// TIA Portal V20 export
FUNCTION_BLOCK "Melden_VisuAllgemein"   // FB127, LAD
{ S7_Optimized_Access := 'TRUE' }
// stored: MemoryReserve 100, SetENOAutomatically false
   VAR
      Register_leer : "Teile Status";
      auf_Seite_Richten { S7_SetPoint := 'True'} : Bool;
      Flanke_Bildwechsel { S7_SetPoint := 'True'} : R_TRIG;
      Bild_tmp { S7_SetPoint := 'True'} : DInt;
      WartezeitSicherung_Reset { S7_SetPoint := 'True'} : TON_TIME;
      Flanke_Türe8_schließen { S7_SetPoint := 'True'} : R_TRIG;
      Flanke_Türe8_öffnen { S7_SetPoint := 'True'} : R_TRIG;
   END_VAR
   VAR RETAIN
      Artikelnummer_tmp { ExternalAccessible := 'False'; ExternalVisible := 'False'; ExternalWritable := 'False'} : String;
   END_VAR
   VAR
      VZ_Leerfahren { S7_SetPoint := 'True'} : TON_TIME;
   END_VAR
   VAR_TEMP
      test : Bool;
   END_VAR
BEGIN

REGION Network 1 (SCL): Richten oder Einzelschrittseite aufgerufen
   CASE "HMI_SYS"."Aktueller Bildschirm" OF
       75:
           #auf_Seite_Richten := true;
       ELSE
           #auf_Seite_Richten := false;
   END_CASE;
END_REGION

REGION Network 2 (SCL): Artikel wurde gewechselt


   IF #Artikelnummer_tmp <> "HMI_COM".Artikelnummer_String THEN
       "HMI_COM".Artikel_gewechselt := true;
       #Artikelnummer_tmp := "HMI_COM".Artikelnummer_String;
   ELSIF "HMI_COM".Grundstellung_Gesamt AND  "HMI_COM".Artikel_gewechselt THEN

       "HMI_COM".Artikel_gewechselt := false;

   END_IF;
END_REGION

NETWORK
TITLE = Übergabe Anwahl Richten
      A     #auf_Seite_Richten;
      JC    m003;

      JU    m001;
m003: NOP   0;

      A     "03_Betriebsart_DB"."NOT-HALT OK";
      A     "03_Betriebsart_DB"."Schutztüren OK";
      JCN   m001;


      A     "HMI_COM".Richten_Gesamtanlage;
      JCN   m002;

      SET;
      S     "HMI_BETR_ART_POS".POS3_0.Taster_Anwahl_GS;


m002: NOP   0;

      A     "HMI_BETR_ART_POS".POS3_0.Taster_Anwahl_GS;
      S     "POS3_0_Signal".Station.SK_Freigabe_Richten;
      =     "POS3_0_Signal".Schrittkette.INIT_SQ;
      R     "HMI_BETR_ART_POS".POS3_0.Taster_Anwahl_GS;


      A     "HMI_COM".Richten_Gesamtanlage;
      R     "HMI_COM".Richten_Gesamtanlage;

m001: NOP   0;


NETWORK
TITLE = Tippbetrieb Aktiv
      A     "POS3_0_Signal".Schrittkette.AUTO_ON;


      =     "HMI_COM".Einzelschritt.Status_Anw;


NETWORK
TITLE = Antriebe sind Ein
      SET;

      =     "HMI_COM".Antriebe_sind_EIN;

REGION Network 6 (SCL): Übergabe Türen Not Halt
   // Allgemeine HMI Übergabe 

   "HMI_COM"."NOT-HALT_OK" := "03_Betriebsart_DB"."NOT-HALT OK";
   "HMI_COM".TUERE_OK := "03_Betriebsart_DB"."Schutztüren OK";




   // Übergabe welche Tür ist nicht verriegelt
   REGION Türen


       "HMI_COM".Tür_offen[1] := "DE_Rueckfuehrung_Tuer_1" AND ("03_Betriebsart_DB".BA_Automatik OR "03_Betriebsart_DB".BA_Manuell OR "03_Betriebsart_DB".BA_Richten);
       "HMI_COM".Tür_offen[2] := "DE_Rueckfuehrung_Tuer_2" AND ("03_Betriebsart_DB".BA_Automatik OR "03_Betriebsart_DB".BA_Manuell OR "03_Betriebsart_DB".BA_Richten);
    //   "HMI_COM".Tür_offen[3] := "DE_Rueckfuehrung_Tuer_3" AND ("03_Betriebsart_DB".BA_Automatik OR "03_Betriebsart_DB".BA_Manuell OR "03_Betriebsart_DB".BA_Richten);
    //   "HMI_COM".Tür_offen[4] := "DE_Rueckfuehrung_Tuer_4" AND ("03_Betriebsart_DB".BA_Automatik OR "03_Betriebsart_DB".BA_Manuell OR "03_Betriebsart_DB".BA_Richten);
    //   "HMI_COM".Tür_offen[5] := "DE_Rueckfuehrung_Tuer_5" AND ("03_Betriebsart_DB".BA_Automatik OR "03_Betriebsart_DB".BA_Manuell OR "03_Betriebsart_DB".BA_Richten);
    //   "HMI_COM".Tür_offen[6] := "DE_Rueckfuehrung_Tuer_6" AND ("03_Betriebsart_DB".BA_Automatik OR "03_Betriebsart_DB".BA_Manuell OR "03_Betriebsart_DB".BA_Richten);
    //   "HMI_COM".Tür_offen[7] := "DE2_0_Rückführung Tür 7" AND ("03_Betriebsart_DB".BA_Automatik OR "03_Betriebsart_DB".BA_Manuell OR "03_Betriebsart_DB".BA_Richten);
    //   "HMI_COM".Tür_offen[8] := "DE2_1_Rückführung Tür 8" AND ("03_Betriebsart_DB".BA_Automatik OR "03_Betriebsart_DB".BA_Manuell OR "03_Betriebsart_DB".BA_Richten);
    (*   "HMI_COM".Tür_offen[9] := "DE2_1_Rückführung Tür 8" AND ("03_Betriebsart_DB".BA_Automatik OR "03_Betriebsart_DB".BA_Manuell OR "03_Betriebsart_DB".BA_Richten);
       "HMI_COM".Tür_offen[10] := "DE2_1_Rückführung Tür 8" AND ("03_Betriebsart_DB".BA_Automatik OR "03_Betriebsart_DB".BA_Manuell OR "03_Betriebsart_DB".BA_Richten);
       "HMI_COM".Tür_offen[11] := "DE2_1_Rückführung Tür 8" AND ("03_Betriebsart_DB".BA_Automatik OR "03_Betriebsart_DB".BA_Manuell OR "03_Betriebsart_DB".BA_Richten);
       "HMI_COM".Tür_offen[12] := "DE2_1_Rückführung Tür 8" AND ("03_Betriebsart_DB".BA_Automatik OR "03_Betriebsart_DB".BA_Manuell OR "03_Betriebsart_DB".BA_Richten);
       "HMI_COM".Tür_offen[13] := "DE2_1_Rückführung Tür 8" AND ("03_Betriebsart_DB".BA_Automatik OR "03_Betriebsart_DB".BA_Manuell OR "03_Betriebsart_DB".BA_Richten);
       "HMI_COM".Tür_offen[14] := "DE2_1_Rückführung Tür 8" AND ("03_Betriebsart_DB".BA_Automatik OR "03_Betriebsart_DB".BA_Manuell OR "03_Betriebsart_DB".BA_Richten);
       "HMI_COM".Tür_offen[15] := "DE2_1_Rückführung Tür 8" AND ("03_Betriebsart_DB".BA_Automatik OR "03_Betriebsart_DB".BA_Manuell OR "03_Betriebsart_DB".BA_Richten); *)
    //   "HMI_COM".Tür_offen[16] := "DE2_1_Rückführung Tür 8" AND ("03_Betriebsart_DB".BA_Automatik OR "03_Betriebsart_DB".BA_Manuell OR "03_Betriebsart_DB".BA_Richten);

   END_REGION
END_REGION

REGION Network 7 (SCL): Rücksetzen der Stationen bei Grundbild



   #Flanke_Bildwechsel(CLK:="03_Betriebsart_DB".BA_Manuell AND #Bild_tmp <> "HMI_SYS"."Aktueller Bildschirm" );



   IF #Flanke_Bildwechsel.Q THEN

       #Bild_tmp := "HMI_SYS"."Aktueller Bildschirm";

    //IF ("HMI_SYS"."Aktueller Bildschirm" = 10125) OR ("03_Betriebsart_DB"."NOT-HALT OK" = false) THEN

       "HMI_COM".Manuell_Zylinder1.Status := 0;
       "HMI_COM".Manuell_Zylinder2.Status := 0;
       "HMI_COM".Manuell_Zylinder3.Status := 0;
       "HMI_COM".Manuell_Zylinder4.Status := 0;

       "HMI_COM".Manuell_Zylinder1.GS := FALSE;
       "HMI_COM".Manuell_Zylinder1.AS1 := FALSE;
       "HMI_COM".Manuell_Zylinder2.GS := FALSE;
       "HMI_COM".Manuell_Zylinder2.AS1 := FALSE;
       "HMI_COM".Manuell_Zylinder3.GS := FALSE;
       "HMI_COM".Manuell_Zylinder3.AS1 := FALSE;
       "HMI_COM".Manuell_Zylinder4.GS := FALSE;
       "HMI_COM".Manuell_Zylinder4.AS1 := FALSE;

      "HMI_COM".Manuell_Zylinder1.DA_GS := FALSE;
       "HMI_COM".Manuell_Zylinder1.DA_AS1 := FALSE;
       "HMI_COM".Manuell_Zylinder2.DA_GS := FALSE;
       "HMI_COM".Manuell_Zylinder2.DA_AS1 := FALSE;
       "HMI_COM".Manuell_Zylinder3.DA_GS := FALSE;
       "HMI_COM".Manuell_Zylinder3.DA_AS1 := FALSE;
       "HMI_COM".Manuell_Zylinder4.DA_GS := FALSE;
       "HMI_COM".Manuell_Zylinder4.DA_AS1 := FALSE;
     END_IF;
END_REGION

REGION Network 8 (SCL): Übertragung und Verwaltung Register



   "HMI_COM".Speichern_Register := false;
END_REGION

REGION Network 9 (SCL): Rucksetzen wenn Register nicht gelöscht
   IF (("HMI_SYS"."Aktueller Bildschirm" = 10001) OR ("HMI_SYS"."Aktueller Bildschirm" = 10010) OR ("HMI_SYS"."Aktueller Bildschirm" = 10020)
       OR ("HMI_SYS"."Aktueller Bildschirm" = 10030)) THEN

       "HMI_BETR_ART_POS".POS3_0.Taster_Reset_Teilestatus := FALSE;
       "HMI_BETR_ART_POS".POS3_1.Taster_Reset_Teilestatus := FALSE;
       "HMI_BETR_ART_POS".POS3_2.Taster_Reset_Teilestatus := FALSE;
       "HMI_BETR_ART_POS".POS3_3.Taster_Reset_Teilestatus := FALSE;
       "HMI_BETR_ART_POS".POS3_4.Taster_Reset_Teilestatus := FALSE;
       "HMI_BETR_ART_POS".POS4_0_Zuführung.Taster_Reset_Teilestatus := FALSE;
       "HMI_BETR_ART_POS".POS5_0_Zuführung.Taster_Reset_Teilestatus := FALSE;
       "HMI_BETR_ART_POS".POS5_0.Taster_Reset_Teilestatus := FALSE;
       "HMI_BETR_ART_POS".POS6_0.Taster_Reset_Teilestatus := FALSE;
       "HMI_BETR_ART_POS".POS7_0.Taster_Reset_Teilestatus := FALSE;
       "HMI_BETR_ART_POS".POS7_1.Taster_Reset_Teilestatus := FALSE;
       "HMI_BETR_ART_POS".POS7_2.Taster_Reset_Teilestatus := FALSE;
       "HMI_BETR_ART_POS".POS7_3.Taster_Reset_Teilestatus := FALSE;
       "HMI_BETR_ART_POS".POS7_4.Taster_Reset_Teilestatus := FALSE;
       "HMI_BETR_ART_POS".POS8_0.Taster_Reset_Teilestatus := FALSE;
       "HMI_BETR_ART_POS".POS9_0.Taster_Reset_Teilestatus := FALSE;
       "HMI_BETR_ART_POS".POS9_1.Taster_Reset_Teilestatus := FALSE;
       "HMI_BETR_ART_POS".POS9_2.Taster_Reset_Teilestatus := FALSE;
       "HMI_BETR_ART_POS".POS9_3.Taster_Reset_Teilestatus := FALSE;
       "HMI_BETR_ART_POS".POS9_4.Taster_Reset_Teilestatus := FALSE;
       "HMI_BETR_ART_POS".POS9_5.Taster_Reset_Teilestatus := FALSE;
       "HMI_BETR_ART_POS".POS9_6.Taster_Reset_Teilestatus := FALSE;
       "HMI_BETR_ART_POS".POS10_0.Taster_Reset_Teilestatus := FALSE;
       "HMI_BETR_ART_POS".POS11.Taster_Reset_Teilestatus := FALSE;
       "HMI_BETR_ART_POS".POS12.Taster_Reset_Teilestatus := FALSE;

   END_IF;
END_REGION

REGION Network 10 (SCL): Leerfahren
   "HMI_Signale".Leerfahren_angewaehlt := "HMI_COM".Leerfahren_angewaehlt;

   #VZ_Leerfahren(IN := "HMI_COM".Leerfahren_ende,
                  PT := t#3s);

   IF #VZ_Leerfahren.Q OR "HMI_COM".Leerfahren_angewaehlt = false THEN

       "HMI_COM".Leerfahren_ende := FALSE;
       "HMI_Signale".Leerfahren_ende := false;
       "HMI_COM".Leerfahren_angewaehlt := false;

       "HMI_COM".Leerfahren_laeuft := false; 
       "POS3_0_Signal".Station.SK_Freigabe_Auto := false;




   END_IF;
END_REGION

REGION Network 11 (SCL): Bildaufrufe


       // Bei Not-Aus Aufruf Grundbild
       IF "03_Betriebsart_DB".BA_0_FP = TRUE OR
           "03_Betriebsart_DB"."NOT-HALT_FN" = TRUE OR
           "03_Betriebsart_DB".Schutztüren_FN = TRUE THEN
           "HMI_SYS".Screen_Name := WSTRING#'B10001_Hauptbild';
       END_IF;


       // Bei BA Manuell Auswahlbild aufrufen
       IF "03_Betriebsart_DB".BA_Manuell_FP = TRUE THEN
           "HMI_SYS".Screen_Name := WSTRING#'B10020_Manuell Auswahl';
       END_IF;


       // Bei BA Richten Auswahlbild aufrufen
       IF "03_Betriebsart_DB".BA_Richten_FP = TRUE THEN
           "HMI_SYS".Screen_Name := WSTRING#'B10075_Übersicht Richten Stationen';
       END_IF;


       // Bei BA Automatik Auswahlbild aufrufen
       IF "03_Betriebsart_DB".BA_Automatik_FP = TRUE THEN
           "HMI_SYS".Screen_Name := WSTRING#'B10010_Automatik';
       END_IF;


       // Bei BA Verwaltung Auswahlbild aufrufen
       IF "03_Betriebsart_DB".BA_Verwaltung_FP = TRUE THEN
           "HMI_SYS".Screen_Name := WSTRING#'B10030_Übersicht Verwaltung';
       END_IF;
END_REGION

REGION Network 12 (SCL): DE +HS1=AN-22T1 Selektivmodul
   #test := NOT "DE_Selektivmodul_OK";

   #WartezeitSicherung_Reset(IN:=#test,
                             PT:=t#25s);





   IF #WartezeitSicherung_Reset.Q = False AND "DE_Selektivmodul_OK"= false THEN
       "HMI_COM".Status_24V_Sicherung := 3;
   ELSIF "DE_Selektivmodul_OK" = false AND "HMI_COM".Status_24V_Sicherung <> 2 THEN
       "HMI_COM".Status_24V_Sicherung  := 0;
   ELSIF "DE_Selektivmodul_OK" = false AND "HMI_COM".Status_24V_Sicherung = 2 THEN
       "DA_Selektivmodul Reset" := true;
   ELSIF "DE_Selektivmodul_OK" THEN
       "HMI_COM".Status_24V_Sicherung := 1;
       "DA_Selektivmodul Reset" := false;
   END_IF;
END_REGION

REGION Network 13 (SCL): nur zum testen
   (* IF "HMI_COM".HMI_Achse_Steuerung.E_jog_pos THEN

       "Pos3_0_Signal".Y_Achse_1.E_jog_pos := true;
       "Pos3_0_Signal".Y_Achse_2.E_jog_pos := true;
       "Pos3_0_Signal".Y_Achse_3.E_jog_pos := true;
       "Pos3_0_Signal".Y_Achse_4.E_jog_pos := true;
       "Pos3_0_Signal".Y_Achse_1.E_jog_neg := 0;
       "Pos3_0_Signal".Y_Achse_2.E_jog_neg := 0;
       "Pos3_0_Signal".Y_Achse_3.E_jog_neg := 0;
       "Pos3_0_Signal".Y_Achse_4.E_jog_neg := 0;

   ELSIF "HMI_COM".HMI_Achse_Steuerung.E_jog_neg THEN


       "Pos3_0_Signal".Y_Achse_1.E_jog_neg := true;
       "Pos3_0_Signal".Y_Achse_2.E_jog_neg := true;
       "Pos3_0_Signal".Y_Achse_3.E_jog_neg := true;
       "Pos3_0_Signal".Y_Achse_4.E_jog_neg := true;

       "Pos3_0_Signal".Y_Achse_1.E_jog_pos := 0;
       "Pos3_0_Signal".Y_Achse_2.E_jog_pos := 0;
       "Pos3_0_Signal".Y_Achse_3.E_jog_pos := 0;
       "Pos3_0_Signal".Y_Achse_4.E_jog_pos := 0;

   ELSE
       "Pos3_0_Signal".Y_Achse_1.E_jog_neg := 0;
       "Pos3_0_Signal".Y_Achse_2.E_jog_neg := 0;
       "Pos3_0_Signal".Y_Achse_3.E_jog_neg := 0;
       "Pos3_0_Signal".Y_Achse_4.E_jog_neg := 0;
       "Pos3_0_Signal".Y_Achse_1.E_jog_pos := 0;
       "Pos3_0_Signal".Y_Achse_2.E_jog_pos := 0;
       "Pos3_0_Signal".Y_Achse_3.E_jog_pos := 0;
       "Pos3_0_Signal".Y_Achse_4.E_jog_pos := 0;
   END_IF; *)

   // "HMI_COM".Manuell_Zylinder1.GS := false;
   // "HMI_COM".Manuell_Zylinder1.AS1 := false;
   // "HMI_COM".Manuell_Zylinder2.GS := false;
   // "HMI_COM".Manuell_Zylinder2.AS1 := false;
   // "HMI_COM".Manuell_Zylinder3.GS := false;
   // "HMI_COM".Manuell_Zylinder3.AS1 := false;
   // "HMI_COM".Manuell_Zylinder4.GS := false;
   // "HMI_COM".Manuell_Zylinder4.AS1 := false;
END_REGION

REGION Network 14 (SCL): Übergabe Taktzeiten Stationen
   "HMI_COM".Taktzeit[0] := "POS3_0_Signal".Taktzeit[0];
END_REGION

REGION Network 15 (SCL): Rücksetzten Messmittelabläufe
   IF ("HMI_COM".Abläufe_Messmittel < 1) OR "03_Betriebsart_DB".Stopp_Taste = false THEN
       "HMI_COM".Messmittel_ein := false;
       ;
   END_IF;


   IF ("HMI_COM".Abläufe_Messmittel_Rundlauf < 1) OR "03_Betriebsart_DB".Stopp_Taste = false THEN
       "HMI_COM".Messmittel_Rundlauf_ein := false;
       ;
   END_IF;
END_REGION
END_FUNCTION_BLOCK
